(* IEC 61131-3 sources: programs/VI-54/VI-54_20171205/VI-54_20171205/Stations/PLC_VI54/VI-54_171014/Class/MyEasy_Filter, 1 file *)

(* ---- MyEasy_Filter.st ---- *)
#include "..\..\Class\MyEasy_Filter\FilterSetting.h"

(*!
<Class
	Name               = "MyEasy_Filter"
	Revision           = "0.0"
	RealtimeTask       = "false"
	CyclicTask         = "true"
	BackgroundTask     = "false"
	Sigmatek           = "false"
	OSInterface        = "false"
	HighPriority       = "false"
	Automatic          = "false"
	UpdateMode         = "Prescan"
	SharedCommandTable = "true"
	Objectsize         = "(480,240)">
	<Channels>
		<Client Name="Div" Required="true" Internal="false"/>
	</Channels>
	<Dependencies>
		<Files>
			<File Path=".\Class\MyEasy_Filter\FilterSetting.h" Include="true"/>
		</Files>
	</Dependencies>
	<Network Name="MyEasy_Filter">
		<!-- List of Components in this network -->
		<Components>
			<Object
				Name       = "_base"
				Class      = "Easy_Filter"
				Position   = "(218,120)"
				Visualized = "true">
				<Channels>
					<Server Name="output"/>
					<Client Name="averages"/>
					<Client Name="input"/>
				</Channels>
			</Object>
		</Components>
		<Comments>
		</Comments>
		<!-- List of Connections in this network -->
		<Connections>
			<Connection Source="this.output" Destination="_base.output" Vertices="(690,210),(518,210),"/>
			<Connection Source="_base.input" Destination="this.input" Vertices="(218,210),(38,210),"/>
			<Connection Source="_base.averages" Destination="this.averages" Vertices="(218,270),(38,270),"/>
		</Connections>
		<!-- Headerfiles -->
		<Options>
		</Options>
	</Network>
</Class>
*)
#pragma using Easy_Filter

MyEasy_Filter : CLASS
: Easy_Filter
  //Servers:
  //Clients:
	Div 	: CltCh_DivEnum;
  //Variables:
		FilterValues : ARRAY [0..Meetingen] OF DINT;

		divide 	: DINT;
  //Functions:
				//! <Function Comment="****************************************************************&#13;&#10;   Easy Digital Filter&#13;&#10;   Filter is only averaging the inputvalue&#13;&#10;****************************************************************&#13;&#10;     Created   :   BS  :   KW46/2001&#13;&#10;****************************************************************&#13;&#10;****************************************************************&#13;&#10;   Einfaches digitales Filter&#13;&#10;   Filter berechnet den Mittelwert der Eingabewerte.&#13;&#10;****************************************************************&#13;&#10;     erstellt  :   BS  :   KW46/2001&#13;&#10;****************************************************************&#13;&#10;" Name="CyWork"/>
	FUNCTION VIRTUAL GLOBAL CyWork
		VAR_INPUT
			EAX 	: UDINT := EAX;
		END_VAR
		VAR_OUTPUT
			state (EAX) 	: UDINT;
		END_VAR;

	FUNCTION GLOBAL Div_Filter
		VAR_OUTPUT
			State 	: DINT;
		END_VAR;
  //Tables:
	FUNCTION @STD
		VAR_OUTPUT
			ret_code	: CONFSTATES;
		END_VAR;
	FUNCTION GLOBAL TAB @CT_;
END_CLASS;

FUNCTION VIRTUAL GLOBAL MyEasy_Filter::CyWork
	VAR_INPUT
		EAX 	: UDINT;
	END_VAR
	VAR_OUTPUT
		state (EAX) 	: UDINT;
	END_VAR

  case Div of
  eDiv1:input   	:= input.read() / 1;
        divide    := 1;
  eDiv10:input   	:= input.read() / 10;
        divide    := 10;
  eDiv100:input 	:= input.read() / 100;
        divide    := 100;
  eDiv1000:input  := input.read() / 1000;
        divide    := 1000;
  else
    div := div.Read();
    divide  := to_dint(Div);
  end_case;

	averages	:= averages.read();

	index_F += 1;

	IF averages <= 0 THEN
		index_F := 0;
	ELSIF index_F >= Averages THEN
		index_F := 0;
		first_full := 1;
	END_IF;

	Sum := Sum - FilterValues[index_F] + input;
	FilterValues[index_F] := input;

	IF averages > 0 & (index_F | first_Full) THEN
		IF averages > Meetingen | averages < 0 THEN
			averages := Meetingen;
        END_IF;
		output := Sum / TO_DINT(averages);
	ELSE
		output := input;
	END_IF;

	state := READY$UDINT;

END_FUNCTION

FUNCTION GLOBAL MyEasy_Filter::Div_Filter
	VAR_OUTPUT
		State 	: DINT;
	END_VAR

  State := Divide;

END_FUNCTION
